PROGRAM MAPPING_in
VAR
  sMapping              : STRING;
  bFirstCycle           : BOOL := TRUE;

  YardState             : U_YARD_STATE;
  TicketListOutput      : U_TICKET_LIST_DATA_OUTPUT;
  TicketListState       : U_TICKET_LIST_STATE;
  InstanceState         : U_INSTANCE_STATE;
  MoverSelectorState    : U_MOVER_SELECTOR_STATE;

  szInstanceState       : ARRAY[1..2] OF UDINT;
  szTicketState         : ARRAY[1..2] OF UDINT;
  szTicketData          : ARRAY[1..2] OF UDINT;
END_VAR


IF (bFirstCycle)
THEN
  bFirstCycle         := FALSE;
  
  szInstanceState[1]  := SIZEOF(InstanceState);
  szInstanceState[2]  := SIZEOF(GVL_APPLICATION.InstanceState);

  szTicketState[1]    := SIZEOF(TicketListState);
  szTicketState[2]    := SIZEOF(GVL_APPLICATION.TicketListState);

  szTicketData[1]     := SIZEOF(TicketListOutput);
  szTicketData[2]     := SIZEOF(GVL_APPLICATION.TicketListDataOutput);
END_IF
//---------------------------------------------------------------------
IF (SIZEOF(TicketListOutput) <> SIZEOF(GVL_APPLICATION.TicketListDataOutput))
THEN
  sMapping  := 'TicketListOutput sizes DO NOT match';
  RETURN;
END_IF
//---------------------------------------------------------------------
IF (SIZEOF(TicketListState) <> SIZEOF(GVL_APPLICATION.TicketListState))
THEN
  sMapping  := 'TicketListState sizes DO NOT match';
  RETURN;
END_IF
//---------------------------------------------------------------------
IF (SIZEOF(InstanceState) <> SIZEOF(GVL_APPLICATION.InstanceState))
THEN
  sMapping  := 'InstanceState sizes DO NOT match';
  RETURN;
END_IF
//---------------------------------------------------------------------
IF (SIZEOF(YardState) <> SIZEOF(GVL_APPLICATION.YardState))
THEN
  sMapping  := 'YardState sizes DO NOT match';
  RETURN;
END_IF
//---------------------------------------------------------------------
IF (SIZEOF(MoverSelectorState) <> SIZEOF(GVL_XTS.MoverSelectorState))
THEN
  sMapping  := 'MoverSelectorState sizes DO NOT match';
  RETURN;
END_IF
//---------------------------------------------------------------------
sMapping    := 'MAPPING ACTIVE';
//-----------------------------------------------------------------------------------------
//       destination,                               source,                   size
//-----------------------------------------------------------------------------------------
  memcpy(ADR(GVL_APPLICATION.YardState),            ADR(YardState),           SIZEOF(YardState));
  memcpy(ADR(GVL_APPLICATION.InstanceState),        ADR(InstanceState),       SIZEOF(InstanceState));
  memcpy(ADR(GVL_APPLICATION.TicketListState),      ADR(TicketListState),     SIZEOF(TicketListState));
  memcpy(ADR(GVL_APPLICATION.TicketListDataOutput), ADR(TicketListOutput),    SIZEOF(TicketListOutput));
  memcpy(ADR(GVL_XTS.MoverSelectorState),           ADR(MoverSelectorState),  SIZEOF(MoverSelectorState));
//-----------------------------------------------------------------------------------------
//-----------------------------------------------------------------------------------------

END_PROGRAM

(* stored: Version 1.1.0.1
   POU MAPPING_in: Id {ebd5c56c-9a35-4de5-bef9-9829dd0bb032}, SpecialFunc None *)
